Fanuc KAREL source: KB00138.KL

PROGRAM KB00138
%NOLOCKGROUP
%ENVIRONMENT CORE
VAR
  P1: STRING[80]
  P2: INTEGER
  P3: INTEGER
BEGIN
  P1 = 'A'
  P2 = 1
  P3 = 1
  PROG_CLEAR(P1, P2, P3)
END KB00138
